// TIA Portal V19 export
// export: Created 2026-10-15T09:44:23.3519815Z, ExportSetting WithDefaults, DisplayName Totally Integrated Automation Portal, DisplayVersion V19, DisplayName TIA Portal Openness, DisplayVersion V19, DisplayName TIA Portal Version Control Interface, DisplayVersion V19, DisplayName STEP 7 Professional, DisplayVersion V19, DisplayName STEP 7 Safety, DisplayVersion V19, DisplayName WinCC Basic/Comfort/Advanced, DisplayVersion V19, DisplayName WinCC Unified, DisplayVersion V19
FUNCTION "ROLL_PB2" : Void   // FC14, SCL
{ S7_Optimized_Access := 'TRUE' }
VERSION : 0.1
// stored: AutoNumber true, IsIECCheckEnabled false, SetENOAutomatically false, UDAEnableTagReadback false
   VAR_TEMP
      r : Bool;
      a1 : Word;
      a2 : Word;
      activeDataBlock : Int;
      comparisonResults : Array[0..0] of Bool;
   END_VAR
BEGIN

   #r := FALSE;
   #a1 := W#16#0000;
   #a2 := W#16#0000;
   #activeDataBlock := 0;
   // PB2, STEP 5 network 1
   #r := ((NOT "ROLL_State".M[0, 1]) AND "ROLL_State".S5Timers[11].Q);
   "ROLL_State".M[4, 1] := #r;
   // PB2, STEP 5 network 2
   #r := ((NOT "ROLL_State".M[4, 1]) OR "ROLL_IO".Input[1, 0]);
   "ROLL_State".M[3, 1] := #r;
   // PB2, STEP 5 network 3
   #r := ((((NOT "ROLL_State".M[31, 4]) AND "ROLL_IO".Input[0, 4] AND "ROLL_State".M[4, 1]) OR "ROLL_State".M[31, 5]) AND "ROLL_IO".Input[0, 2]);
   "ROLL_State".M[4, 4] := #r;
   // PB2, STEP 5 network 4
   #r := (NOT "ROLL_IO".Input[11, 7]);
   IF #r THEN
       "ROLL_State".M[5, 0] := TRUE;
   END_IF;
   #r := "ROLL_State".M[3, 1];
   IF #r THEN
       "ROLL_State".M[5, 0] := FALSE;
   END_IF;
   // PB2, STEP 5 network 5
   #r := (NOT "ROLL_IO".Input[13, 5]);
   IF #r THEN
       "ROLL_State".M[5, 1] := TRUE;
   END_IF;
   #r := "ROLL_State".M[3, 1];
   IF #r THEN
       "ROLL_State".M[5, 1] := FALSE;
   END_IF;
   // PB2, STEP 5 network 6
   #r := (NOT "ROLL_IO".Input[13, 0]);
   IF #r THEN
       "ROLL_State".M[5, 2] := TRUE;
   END_IF;
   #r := "ROLL_State".M[3, 1];
   IF #r THEN
       "ROLL_State".M[5, 2] := FALSE;
   END_IF;
   // PB2, STEP 5 network 7
   #r := (NOT "ROLL_IO".Input[8, 5]);
   IF #r THEN
       "ROLL_State".M[5, 3] := TRUE;
   END_IF;
   #r := "ROLL_State".M[3, 1];
   IF #r THEN
       "ROLL_State".M[5, 3] := FALSE;
   END_IF;
   // PB2, STEP 5 network 8
   #r := "ROLL_State".M[0, 3];
   IF #r THEN
       "ROLL_State".M[5, 4] := TRUE;
   END_IF;
   #r := "ROLL_State".M[3, 1];
   IF #r THEN
       "ROLL_State".M[5, 4] := FALSE;
   END_IF;
   // PB2, STEP 5 network 9
   #r := "ROLL_State".M[0, 3];
   IF #r THEN
       "ROLL_State".M[5, 5] := TRUE;
   END_IF;
   #r := "ROLL_State".M[3, 1];
   IF #r THEN
       "ROLL_State".M[5, 5] := FALSE;
   END_IF;
   // PB2, STEP 5 network 10
   #r := "ROLL_IO".Input[3, 6];
   IF #r THEN
       "ROLL_State".M[5, 6] := TRUE;
   END_IF;
   #r := "ROLL_State".M[3, 1];
   IF #r THEN
       "ROLL_State".M[5, 6] := FALSE;
   END_IF;
   // PB2, STEP 5 network 11
   #r := (NOT "ROLL_IO".Input[3, 7]);
   IF #r THEN
       "ROLL_State".M[5, 7] := TRUE;
   END_IF;
   #r := "ROLL_State".M[3, 1];
   IF #r THEN
       "ROLL_State".M[5, 7] := FALSE;
   END_IF;
   // PB2, STEP 5 network 12
   #r := (NOT "ROLL_IO".Input[5, 2]);
   IF #r THEN
       "ROLL_State".M[6, 0] := TRUE;
   END_IF;
   #r := ("ROLL_IO".Input[5, 2] AND "ROLL_State".M[3, 1]);
   IF #r THEN
       "ROLL_State".M[6, 0] := FALSE;
   END_IF;
   // PB2, STEP 5 network 13
   #r := ((NOT "ROLL_IO".Input[5, 3]) AND "ROLL_State".S5Timers[31].Q);
   IF #r THEN
       "ROLL_State".M[6, 1] := TRUE;
   END_IF;
   #r := "ROLL_State".M[3, 1];
   IF #r THEN
       "ROLL_State".M[6, 1] := FALSE;
   END_IF;
   // PB2, STEP 5 network 14
   #r := (NOT "ROLL_IO".Input[5, 4]);
   IF #r THEN
       "ROLL_State".M[6, 2] := TRUE;
   END_IF;
   #r := ("ROLL_IO".Input[5, 4] AND "ROLL_State".M[3, 1]);
   IF #r THEN
       "ROLL_State".M[6, 2] := FALSE;
   END_IF;
   // PB2, STEP 5 network 15
   #r := ((NOT "ROLL_IO".Input[5, 5]) AND "ROLL_State".M[40, 5] AND "ROLL_State".S5Timers[17].Q);
   IF #r THEN
       "ROLL_State".M[6, 3] := TRUE;
   END_IF;
   #r := "ROLL_State".M[3, 1];
   IF #r THEN
       "ROLL_State".M[6, 3] := FALSE;
   END_IF;
   // PB2, STEP 5 network 16
   #r := ((NOT "ROLL_IO".Input[6, 0]) AND "ROLL_State".S5Timers[32].Q);
   IF #r THEN
       "ROLL_State".M[6, 4] := TRUE;
   END_IF;
   #r := "ROLL_State".M[3, 1];
   IF #r THEN
       "ROLL_State".M[6, 4] := FALSE;
   END_IF;
   // PB2, STEP 5 network 17
   #r := ((NOT "ROLL_IO".Input[6, 2]) AND "ROLL_State".S5Timers[33].Q);
   IF #r THEN
       "ROLL_State".M[6, 5] := TRUE;
   END_IF;
   #r := "ROLL_State".M[3, 1];
   IF #r THEN
       "ROLL_State".M[6, 5] := FALSE;
   END_IF;
   // PB2, STEP 5 network 18
   #r := "ROLL_State".M[0, 3];
   IF #r THEN
       "ROLL_State".M[6, 6] := TRUE;
   END_IF;
   #r := "ROLL_State".M[3, 1];
   IF #r THEN
       "ROLL_State".M[6, 6] := FALSE;
   END_IF;
   // PB2, STEP 5 network 19
   #r := ((NOT "ROLL_State".M[0, 3]) AND "ROLL_State".S5Timers[35].Q);
   IF #r THEN
       "ROLL_State".M[6, 7] := TRUE;
   END_IF;
   #r := "ROLL_State".M[3, 1];
   IF #r THEN
       "ROLL_State".M[6, 7] := FALSE;
   END_IF;
   // PB2, STEP 5 network 20
   #r := ((NOT "ROLL_State".M[0, 3]) AND "ROLL_State".S5Timers[36].Q);
   IF #r THEN
       "ROLL_State".M[7, 0] := TRUE;
   END_IF;
   #r := "ROLL_State".M[3, 1];
   IF #r THEN
       "ROLL_State".M[7, 0] := FALSE;
   END_IF;
   // PB2, STEP 5 network 21
   #r := ((NOT "ROLL_State".M[0, 3]) AND "ROLL_State".M[48, 1] AND "ROLL_State".S5Timers[37].Q);
   IF #r THEN
       "ROLL_State".M[7, 1] := TRUE;
   END_IF;
   #r := "ROLL_State".M[3, 1];
   IF #r THEN
       "ROLL_State".M[7, 1] := FALSE;
   END_IF;
   // PB2, STEP 5 network 22
   #r := ((NOT "ROLL_State".M[0, 3]) AND "ROLL_State".S5Timers[38].Q);
   IF #r THEN
       "ROLL_State".M[7, 2] := TRUE;
   END_IF;
   #r := "ROLL_State".M[3, 1];
   IF #r THEN
       "ROLL_State".M[7, 2] := FALSE;
   END_IF;
   // PB2, STEP 5 network 23
   #r := ((NOT "ROLL_IO".Input[5, 6]) AND "ROLL_State".S5Timers[16].Q);
   IF #r THEN
       "ROLL_State".M[7, 3] := TRUE;
   END_IF;
   #r := ("ROLL_IO".Input[5, 6] AND "ROLL_State".M[3, 1]);
   IF #r THEN
       "ROLL_State".M[7, 3] := FALSE;
   END_IF;
   // PB2, STEP 5 network 24
   #r := "ROLL_State".M[0, 3];
   IF #r THEN
       "ROLL_State".M[7, 4] := TRUE;
   END_IF;
   #r := "ROLL_State".M[3, 1];
   IF #r THEN
       "ROLL_State".M[7, 4] := FALSE;
   END_IF;
   // PB2, STEP 5 network 25
   #r := "ROLL_State".M[0, 3];
   IF #r THEN
       "ROLL_State".M[7, 5] := TRUE;
   END_IF;
   #r := "ROLL_State".M[3, 1];
   IF #r THEN
       "ROLL_State".M[7, 5] := FALSE;
   END_IF;
   // PB2, STEP 5 network 26
   #r := "ROLL_State".M[0, 3];
   IF #r THEN
       "ROLL_State".M[7, 6] := TRUE;
   END_IF;
   #r := "ROLL_State".M[3, 1];
   IF #r THEN
       "ROLL_State".M[7, 6] := FALSE;
   END_IF;
   // PB2, STEP 5 network 27
   #r := (NOT "ROLL_IO".Input[6, 7]);
   IF #r THEN
       "ROLL_State".M[7, 7] := TRUE;
   END_IF;
   #r := "ROLL_State".M[3, 1];
   IF #r THEN
       "ROLL_State".M[7, 7] := FALSE;
   END_IF;
   // PB2, STEP 5 network 28
   #a2 := #a1;
   #a1 := W#16#1050;
   #r := ((NOT "ROLL_IO".Input[7, 6]) AND "ROLL_IO".Output[20, 5]);
   "ROLL_TimerOp"(Number := 30,
                  Operation := 0,
                  Signal := #r,
                  Preset := #a1);
   #r := "ROLL_State".S5Timers[30].Q;
   IF #r THEN
       "ROLL_State".M[8, 6] := TRUE;
   END_IF;
   #r := "ROLL_State".M[3, 1];
   IF #r THEN
       "ROLL_State".M[8, 6] := FALSE;
   END_IF;
   // PB2, STEP 5 network 29
   #r := "ROLL_State".M[0, 3];
   IF #r THEN
       "ROLL_State".M[8, 7] := TRUE;
   END_IF;
   #r := "ROLL_State".M[3, 1];
   IF #r THEN
       "ROLL_State".M[8, 7] := FALSE;
   END_IF;
   // PB2, STEP 5 network 30
   #r := ((NOT "ROLL_IO".Input[13, 7]) AND "ROLL_State".M[4, 1]);
   IF #r THEN
       "ROLL_State".M[9, 0] := TRUE;
   END_IF;
   #r := ("ROLL_IO".Input[13, 7] AND "ROLL_State".M[3, 1]);
   IF #r THEN
       "ROLL_State".M[9, 0] := FALSE;
   END_IF;
   // PB2, STEP 5 network 31
   #r := "ROLL_State".M[0, 3];
   IF #r THEN
       "ROLL_State".M[9, 1] := TRUE;
   END_IF;
   #r := "ROLL_State".M[3, 1];
   IF #r THEN
       "ROLL_State".M[9, 1] := FALSE;
   END_IF;
   // PB2, STEP 5 network 32
   #r := ((NOT "ROLL_State".M[28, 4]) AND (NOT "ROLL_State".M[31, 5]) AND (((NOT "ROLL_State".M[20, 2]) AND ("ROLL_IO".Input[123, 5] OR "ROLL_IO".Input[123, 6])) OR "ROLL_State".M[70, 2] OR "ROLL_State".M[70, 3]) AND "ROLL_IO".Input[0, 4] AND "ROLL_State".M[4, 1]);
   IF #r THEN
       "ROLL_State".M[9, 2] := TRUE;
   END_IF;
   #r := "ROLL_State".M[3, 1];
   IF #r THEN
       "ROLL_State".M[9, 2] := FALSE;
   END_IF;
   // PB2, STEP 5 network 33
   #r := ("ROLL_State".M[4, 1] AND "ROLL_State".S5Timers[19].Q);
   IF #r THEN
       "ROLL_State".M[9, 3] := TRUE;
   END_IF;
   #r := "ROLL_State".M[3, 1];
   IF #r THEN
       "ROLL_State".M[9, 3] := FALSE;
   END_IF;
   // PB2, STEP 5 network 34
   #r := (((("ROLL_State".M[20, 4] OR "ROLL_State".M[20, 5]) AND "ROLL_IO".Input[0, 1] AND "ROLL_State".M[190, 6]) OR "ROLL_State".M[31, 5]) AND "ROLL_State".S5Timers[95].Q);
   "ROLL_State".M[9, 4] := #r;
   // PB2, STEP 5 network 35
   #r := "ROLL_State".M[0, 3];
   IF #r THEN
       "ROLL_State".M[9, 5] := TRUE;
   END_IF;
   #r := "ROLL_State".M[3, 1];
   IF #r THEN
       "ROLL_State".M[9, 5] := FALSE;
   END_IF;
   // PB2, STEP 5 network 36
   #r := "ROLL_State".M[0, 3];
   IF #r THEN
       "ROLL_State".M[9, 6] := TRUE;
   END_IF;
   #r := "ROLL_State".M[3, 1];
   IF #r THEN
       "ROLL_State".M[9, 6] := FALSE;
   END_IF;
   // PB2, STEP 5 network 37
   #r := "ROLL_State".M[0, 3];
   IF #r THEN
       "ROLL_State".M[9, 7] := TRUE;
   END_IF;
   #r := "ROLL_State".M[3, 1];
   IF #r THEN
       "ROLL_State".M[9, 7] := FALSE;
   END_IF;
   // PB2, STEP 5 network 38
   #r := ((NOT "ROLL_IO".Input[12, 0]) AND "ROLL_State".M[4, 1]);
   IF #r THEN
       "ROLL_State".M[10, 0] := TRUE;
   END_IF;
   #r := (((((NOT "ROLL_State".S5Timers[11].Q) AND "ROLL_IO".Input[3, 0]) OR "ROLL_IO".Input[12, 5]) AND "ROLL_State".M[3, 1]) OR (NOT "ROLL_State".M[4, 1]) OR "ROLL_State".M[0, 7]);
   IF #r THEN
       "ROLL_State".M[10, 0] := FALSE;
   END_IF;
   // PB2, STEP 5 network 39
   #r := ((NOT "ROLL_IO".Input[12, 6]) AND "ROLL_State".M[4, 1]);
   IF #r THEN
       "ROLL_State".M[10, 1] := TRUE;
   END_IF;
   #r := (((((NOT "ROLL_State".S5Timers[11].Q) AND "ROLL_IO".Input[3, 0]) OR "ROLL_IO".Input[12, 1]) AND "ROLL_State".M[3, 1]) OR (NOT "ROLL_State".M[4, 1]) OR "ROLL_State".M[0, 7]);
   IF #r THEN
       "ROLL_State".M[10, 1] := FALSE;
   END_IF;
   // PB2, STEP 5 network 40
   #r := "ROLL_State".M[0, 3];
   IF #r THEN
       "ROLL_State".M[10, 2] := TRUE;
   END_IF;
   #r := "ROLL_State".M[3, 1];
   IF #r THEN
       "ROLL_State".M[10, 2] := FALSE;
   END_IF;
   // PB2, STEP 5 network 41
   #r := "ROLL_State".M[0, 3];
   IF #r THEN
       "ROLL_State".M[10, 3] := TRUE;
   END_IF;
   #r := "ROLL_State".M[3, 1];
   IF #r THEN
       "ROLL_State".M[10, 3] := FALSE;
   END_IF;
   // PB2, STEP 5 network 42
   #r := "ROLL_State".M[0, 3];
   IF #r THEN
       "ROLL_State".M[10, 4] := TRUE;
   END_IF;
   #r := "ROLL_State".M[3, 1];
   IF #r THEN
       "ROLL_State".M[10, 4] := FALSE;
   END_IF;
   // PB2, STEP 5 network 43
   #r := "ROLL_State".M[0, 3];
   IF #r THEN
       "ROLL_State".M[10, 5] := TRUE;
   END_IF;
   #r := "ROLL_State".M[3, 1];
   IF #r THEN
       "ROLL_State".M[10, 5] := FALSE;
   END_IF;
   // PB2, STEP 5 network 44
   #r := "ROLL_State".M[0, 3];
   IF #r THEN
       "ROLL_State".M[10, 6] := TRUE;
   END_IF;
   #r := "ROLL_State".M[3, 1];
   IF #r THEN
       "ROLL_State".M[10, 6] := FALSE;
   END_IF;
   // PB2, STEP 5 network 45
   #r := "ROLL_State".M[0, 3];
   IF #r THEN
       "ROLL_State".M[10, 7] := TRUE;
   END_IF;
   #r := "ROLL_State".M[3, 1];
   IF #r THEN
       "ROLL_State".M[10, 7] := FALSE;
   END_IF;
   // PB2, STEP 5 network 46
   #r := ("ROLL_State".M[4, 1] AND "ROLL_State".M[63, 2]);
   IF #r THEN
       "ROLL_State".M[11, 0] := TRUE;
   END_IF;
   #r := "ROLL_State".M[3, 1];
   IF #r THEN
       "ROLL_State".M[11, 0] := FALSE;
   END_IF;
   // PB2, STEP 5 network 47
   #r := ("ROLL_IO".Input[13, 3] AND "ROLL_State".M[4, 1] AND "ROLL_State".S5Timers[112].Q);
   IF #r THEN
       "ROLL_State".M[11, 1] := TRUE;
   END_IF;
   #r := "ROLL_State".M[3, 1];
   IF #r THEN
       "ROLL_State".M[11, 1] := FALSE;
   END_IF;
   // PB2, STEP 5 network 48
   #r := ((NOT "ROLL_IO".Input[13, 3]) AND "ROLL_State".M[4, 1] AND "ROLL_State".S5Timers[15].Q);
   IF #r THEN
       "ROLL_State".M[11, 2] := TRUE;
   END_IF;
   #r := "ROLL_State".M[3, 1];
   IF #r THEN
       "ROLL_State".M[11, 2] := FALSE;
   END_IF;
   // PB2, STEP 5 network 49
   #r := ("ROLL_State".M[4, 1] AND "ROLL_State".M[63, 3]);
   IF #r THEN
       "ROLL_State".M[11, 3] := TRUE;
   END_IF;
   #r := "ROLL_State".M[3, 1];
   IF #r THEN
       "ROLL_State".M[11, 3] := FALSE;
   END_IF;
   // PB2, STEP 5 network 50
   #r := ("ROLL_State".M[190, 6] AND "ROLL_State".M[23, 2] AND "ROLL_State".M[60, 3]);
   IF #r THEN
       "ROLL_State".M[11, 4] := TRUE;
   END_IF;
   #r := "ROLL_State".M[3, 1];
   IF #r THEN
       "ROLL_State".M[11, 4] := FALSE;
   END_IF;
   // PB2, STEP 5 network 51
   #r := "ROLL_State".M[0, 3];
   IF #r THEN
       "ROLL_State".M[11, 5] := TRUE;
   END_IF;
   #r := "ROLL_State".M[3, 1];
   IF #r THEN
       "ROLL_State".M[11, 5] := FALSE;
   END_IF;
   // PB2, STEP 5 network 52
   #r := "ROLL_State".M[0, 3];
   IF #r THEN
       "ROLL_State".M[11, 6] := TRUE;
   END_IF;
   #r := "ROLL_State".M[3, 1];
   IF #r THEN
       "ROLL_State".M[11, 6] := FALSE;
   END_IF;
   // PB2, STEP 5 network 53
   #r := "ROLL_State".M[0, 3];
   IF #r THEN
       "ROLL_State".M[11, 7] := TRUE;
   END_IF;
   #r := "ROLL_State".M[3, 1];
   IF #r THEN
       "ROLL_State".M[11, 7] := FALSE;
   END_IF;
   // PB2, STEP 5 network 54
   #r := (NOT "ROLL_IO".Input[8, 3]);
   IF #r THEN
       "ROLL_State".M[12, 0] := TRUE;
   END_IF;
   #r := "ROLL_State".M[3, 1];
   IF #r THEN
       "ROLL_State".M[12, 0] := FALSE;
   END_IF;
   // PB2, STEP 5 network 55
   #r := ((NOT "ROLL_IO".Input[0, 7]) AND (NOT "ROLL_IO".Input[1, 4]) AND "ROLL_State".M[4, 4]);
   IF #r THEN
       "ROLL_State".M[12, 1] := TRUE;
   END_IF;
   #r := "ROLL_State".M[3, 1];
   IF #r THEN
       "ROLL_State".M[12, 1] := FALSE;
   END_IF;
   // PB2, STEP 5 network 56
   #r := "ROLL_State".M[0, 3];
   IF #r THEN
       "ROLL_State".M[12, 2] := TRUE;
   END_IF;
   #r := "ROLL_State".M[3, 1];
   IF #r THEN
       "ROLL_State".M[12, 2] := FALSE;
   END_IF;
   // PB2, STEP 5 network 57
   #r := "ROLL_State".M[0, 3];
   IF #r THEN
       "ROLL_State".M[12, 3] := TRUE;
   END_IF;
   #r := "ROLL_State".M[3, 1];
   IF #r THEN
       "ROLL_State".M[12, 3] := FALSE;
   END_IF;
   // PB2, STEP 5 network 58
   #r := "ROLL_State".M[0, 3];
   IF #r THEN
       "ROLL_State".M[13, 0] := TRUE;
   END_IF;
   #r := "ROLL_State".M[3, 1];
   IF #r THEN
       "ROLL_State".M[13, 0] := FALSE;
   END_IF;
   // PB2, STEP 5 network 59
   #r := (NOT "ROLL_IO".Input[3, 2]);
   IF #r THEN
       "ROLL_State".M[13, 1] := TRUE;
   END_IF;
   #r := "ROLL_State".M[3, 1];
   IF #r THEN
       "ROLL_State".M[13, 1] := FALSE;
   END_IF;
   // PB2, STEP 5 network 60
   #r := ((NOT "ROLL_IO".Input[4, 7]) AND "ROLL_IO".Input[0, 1] AND "ROLL_State".M[190, 6] AND "ROLL_State".M[27, 4]);
   IF #r THEN
       "ROLL_State".M[13, 2] := TRUE;
   END_IF;
   #r := "ROLL_State".M[3, 1];
   IF #r THEN
       "ROLL_State".M[13, 2] := FALSE;
   END_IF;
   // PB2, STEP 5 network 61
   #r := (NOT "ROLL_IO".Input[5, 0]);
   IF #r THEN
       "ROLL_State".M[13, 3] := TRUE;
   END_IF;
   #r := ("ROLL_IO".Input[5, 0] AND "ROLL_State".M[3, 1]);
   IF #r THEN
       "ROLL_State".M[13, 3] := FALSE;
   END_IF;
   // PB2, STEP 5 network 62
   #r := (NOT "ROLL_IO".Input[10, 7]);
   IF #r THEN
       "ROLL_State".M[13, 4] := TRUE;
   END_IF;
   #r := ("ROLL_IO".Input[10, 7] AND "ROLL_State".M[3, 1]);
   IF #r THEN
       "ROLL_State".M[13, 4] := FALSE;
   END_IF;
   // PB2, STEP 5 network 63
   #r := (NOT "ROLL_IO".Input[4, 5]);
   IF #r THEN
       "ROLL_State".M[13, 7] := TRUE;
   END_IF;
   #r := "ROLL_State".M[3, 1];
   IF #r THEN
       "ROLL_State".M[13, 7] := FALSE;
   END_IF;
   // PB2, STEP 5 network 64
   #a2 := #a1;
   #a1 := W#16#2020;
   #r := (((NOT "ROLL_IO".Input[10, 0]) OR (NOT "ROLL_IO".Input[10, 1]) OR (NOT "ROLL_IO".Input[10, 2]) OR (NOT "ROLL_IO".Input[10, 3])) AND "ROLL_IO".Output[19, 1]);
   "ROLL_TimerOp"(Number := 50,
                  Operation := 0,
                  Signal := #r,
                  Preset := #a1);
   // PB2, STEP 5 network 65
   #r := ((NOT "ROLL_IO".Input[10, 0]) AND "ROLL_State".S5Timers[50].Q);
   IF #r THEN
       "ROLL_State".M[14, 0] := TRUE;
   END_IF;
   #r := "ROLL_State".M[3, 1];
   IF #r THEN
       "ROLL_State".M[14, 0] := FALSE;
   END_IF;
   // PB2, STEP 5 network 66
   #r := ((NOT "ROLL_IO".Input[10, 1]) AND "ROLL_State".S5Timers[50].Q);
   IF #r THEN
       "ROLL_State".M[14, 1] := TRUE;
   END_IF;
   #r := "ROLL_State".M[3, 1];
   IF #r THEN
       "ROLL_State".M[14, 1] := FALSE;
   END_IF;
   // PB2, STEP 5 network 67
   #r := ((NOT "ROLL_IO".Input[10, 2]) AND "ROLL_State".S5Timers[50].Q);
   IF #r THEN
       "ROLL_State".M[14, 2] := TRUE;
   END_IF;
   #r := "ROLL_State".M[3, 1];
   IF #r THEN
       "ROLL_State".M[14, 2] := FALSE;
   END_IF;
   // PB2, STEP 5 network 68
   #r := ((NOT "ROLL_IO".Input[10, 3]) AND "ROLL_State".S5Timers[50].Q);
   IF #r THEN
       "ROLL_State".M[14, 3] := TRUE;
   END_IF;
   #r := "ROLL_State".M[3, 1];
   IF #r THEN
       "ROLL_State".M[14, 3] := FALSE;
   END_IF;
   // PB2, STEP 5 network 69
   #r := "ROLL_State".M[0, 3];
   IF #r THEN
       "ROLL_State".M[15, 2] := TRUE;
   END_IF;
   #r := "ROLL_State".M[3, 1];
   IF #r THEN
       "ROLL_State".M[15, 2] := FALSE;
   END_IF;
   // PB2, STEP 5 network 70
   #r := "ROLL_State".M[0, 3];
   IF #r THEN
       "ROLL_State".M[15, 3] := TRUE;
   END_IF;
   #r := "ROLL_State".M[3, 1];
   IF #r THEN
       "ROLL_State".M[15, 3] := FALSE;
   END_IF;
   // PB2, STEP 5 network 71
   #r := "ROLL_State".M[0, 3];
   IF #r THEN
       "ROLL_State".M[15, 4] := TRUE;
   END_IF;
   #r := "ROLL_State".M[3, 1];
   IF #r THEN
       "ROLL_State".M[15, 4] := FALSE;
   END_IF;
   // PB2, STEP 5 network 72
   #r := (NOT "ROLL_IO".Input[4, 0]);
   IF #r THEN
       "ROLL_State".M[15, 5] := TRUE;
   END_IF;
   #r := "ROLL_State".M[3, 1];
   IF #r THEN
       "ROLL_State".M[15, 5] := FALSE;
   END_IF;
   // PB2, STEP 5 network 73
   #r := (NOT "ROLL_IO".Input[4, 1]);
   IF #r THEN
       "ROLL_State".M[15, 6] := TRUE;
   END_IF;
   #r := "ROLL_State".M[3, 1];
   IF #r THEN
       "ROLL_State".M[15, 6] := FALSE;
   END_IF;
   // PB2, STEP 5 network 74
   #r := (NOT "ROLL_IO".Input[4, 2]);
   IF #r THEN
       "ROLL_State".M[15, 7] := TRUE;
   END_IF;
   #r := "ROLL_State".M[3, 1];
   IF #r THEN
       "ROLL_State".M[15, 7] := FALSE;
   END_IF;
   // PB2, STEP 5 network 75
   #r := "ROLL_State".M[16, 0];
   IF #r THEN
       "ROLL_State".M[16, 0] := TRUE;
   END_IF;
   #r := "ROLL_State".M[3, 1];
   IF #r THEN
       "ROLL_State".M[16, 0] := FALSE;
   END_IF;
   // PB2, STEP 5 network 76
   #r := "ROLL_State".M[16, 1];
   IF #r THEN
       "ROLL_State".M[16, 1] := TRUE;
   END_IF;
   #r := "ROLL_State".M[3, 1];
   IF #r THEN
       "ROLL_State".M[16, 1] := FALSE;
   END_IF;
   // PB2, STEP 5 network 77
   #r := "ROLL_State".M[16, 2];
   IF #r THEN
       "ROLL_State".M[16, 2] := TRUE;
   END_IF;
   #r := "ROLL_State".M[3, 1];
   IF #r THEN
       "ROLL_State".M[16, 2] := FALSE;
   END_IF;
   // PB2, STEP 5 network 78
   #r := ("ROLL_State".M[34, 1] AND "ROLL_State".M[4, 1]);
   IF #r THEN
       "ROLL_State".M[16, 3] := TRUE;
   END_IF;
   #r := "ROLL_State".M[3, 1];
   IF #r THEN
       "ROLL_State".M[16, 3] := FALSE;
   END_IF;
   // PB2, STEP 5 network 79
   #r := "ROLL_State".M[16, 4];
   IF #r THEN
       "ROLL_State".M[16, 4] := TRUE;
   END_IF;
   #r := ((NOT "ROLL_IO".Input[123, 1]) AND (NOT "ROLL_IO".Input[123, 4]) AND (NOT "ROLL_IO".Input[123, 5]) AND (NOT "ROLL_IO".Input[123, 6]) AND (NOT "ROLL_IO".Input[125, 0]) AND (NOT "ROLL_IO".Input[125, 1]) AND "ROLL_State".M[3, 1]);
   IF #r THEN
       "ROLL_State".M[16, 4] := FALSE;
   END_IF;
   // PB2, STEP 5 network 80
   #r := "ROLL_State".M[16, 5];
   IF #r THEN
       "ROLL_State".M[16, 5] := TRUE;
   END_IF;
   #r := "ROLL_State".M[3, 1];
   IF #r THEN
       "ROLL_State".M[16, 5] := FALSE;
   END_IF;
   // PB2, STEP 5 network 81
   #r := ((NOT "ROLL_IO".Input[3, 4]) AND "ROLL_State".M[4, 1]);
   IF #r THEN
       "ROLL_State".M[16, 6] := TRUE;
   END_IF;
   #r := ("ROLL_IO".Input[3, 4] AND "ROLL_State".M[3, 1]);
   IF #r THEN
       "ROLL_State".M[16, 6] := FALSE;
   END_IF;
   // PB2, STEP 5 network 82
   #r := ((NOT "ROLL_IO".Input[3, 1]) AND ((("ROLL_State".M[190, 5] OR "ROLL_State".M[190, 6]) AND "ROLL_IO".Input[0, 1]) OR "ROLL_State".M[4, 4]) AND "ROLL_State".M[4, 1]);
   IF #r THEN
       "ROLL_State".M[16, 7] := TRUE;
   END_IF;
   #r := "ROLL_State".M[3, 1];
   IF #r THEN
       "ROLL_State".M[16, 7] := FALSE;
   END_IF;
   // PB2, STEP 5 network 83
   #r := ((NOT "ROLL_IO".Input[3, 5]) AND "ROLL_State".M[4, 1]);
   IF #r THEN
       "ROLL_State".M[17, 0] := TRUE;
   END_IF;
   #r := ("ROLL_IO".Input[3, 5] AND "ROLL_State".M[3, 1]);
   IF #r THEN
       "ROLL_State".M[17, 0] := FALSE;
   END_IF;
   // PB2, STEP 5 network 84
   #r := "ROLL_State".M[0, 3];
   IF #r THEN
       "ROLL_State".M[17, 1] := TRUE;
   END_IF;
   #r := "ROLL_State".M[3, 1];
   IF #r THEN
       "ROLL_State".M[17, 1] := FALSE;
   END_IF;
   // PB2, STEP 5 network 85
   #r := "ROLL_State".M[0, 3];
   IF #r THEN
       "ROLL_State".M[17, 2] := TRUE;
   END_IF;
   #r := "ROLL_State".M[3, 1];
   IF #r THEN
       "ROLL_State".M[17, 2] := FALSE;
   END_IF;
   // PB2, STEP 5 network 86
   #r := "ROLL_State".M[0, 3];
   IF #r THEN
       "ROLL_State".M[17, 3] := TRUE;
   END_IF;
   #r := "ROLL_State".M[3, 1];
   IF #r THEN
       "ROLL_State".M[17, 3] := FALSE;
   END_IF;
   // PB2, STEP 5 network 87
   #r := "ROLL_State".M[0, 3];
   IF #r THEN
       "ROLL_State".M[17, 4] := TRUE;
   END_IF;
   #r := "ROLL_State".M[3, 1];
   IF #r THEN
       "ROLL_State".M[17, 4] := FALSE;
   END_IF;
   // PB2, STEP 5 network 88
   #r := "ROLL_State".M[0, 3];
   IF #r THEN
       "ROLL_State".M[17, 5] := TRUE;
   END_IF;
   #r := "ROLL_State".M[3, 1];
   IF #r THEN
       "ROLL_State".M[17, 5] := FALSE;
   END_IF;
   // PB2, STEP 5 network 89
   #r := "ROLL_State".M[0, 3];
   IF #r THEN
       "ROLL_State".M[17, 6] := TRUE;
   END_IF;
   #r := "ROLL_State".M[3, 1];
   IF #r THEN
       "ROLL_State".M[17, 6] := FALSE;
   END_IF;
   // PB2, STEP 5 network 90
   #r := "ROLL_State".M[0, 3];
   IF #r THEN
       "ROLL_State".M[17, 7] := TRUE;
   END_IF;
   #r := "ROLL_State".M[3, 1];
   IF #r THEN
       "ROLL_State".M[17, 7] := FALSE;
   END_IF;
   // PB2, STEP 5 network 91
   #r := "ROLL_State".M[0, 3];
   IF #r THEN
       "ROLL_State".M[18, 0] := TRUE;
   END_IF;
   #r := "ROLL_State".M[3, 1];
   IF #r THEN
       "ROLL_State".M[18, 0] := FALSE;
   END_IF;
   // PB2, STEP 5 network 92
   #r := ((NOT "ROLL_IO".Input[14, 0]) AND ((("ROLL_State".M[190, 5] OR "ROLL_State".M[190, 6]) AND ("ROLL_State".M[23, 0] OR "ROLL_State".M[23, 1] OR "ROLL_State".M[23, 2] OR "ROLL_State".M[23, 3])) OR ("ROLL_State".M[16, 3] AND "ROLL_State".M[31, 4] AND "ROLL_State".M[37, 2]) OR "ROLL_State".M[74, 0]));
   IF #r THEN
       "ROLL_State".M[18, 1] := TRUE;
   END_IF;
   #r := "ROLL_State".M[3, 1];
   IF #r THEN
       "ROLL_State".M[18, 1] := FALSE;
   END_IF;
   // PB2, STEP 5 network 93
   #r := "ROLL_State".M[0, 3];
   IF #r THEN
       "ROLL_State".M[18, 2] := TRUE;
   END_IF;
   #r := "ROLL_State".M[3, 1];
   IF #r THEN
       "ROLL_State".M[18, 2] := FALSE;
   END_IF;
   // PB2, STEP 5 network 94
   #r := "ROLL_State".M[0, 3];
   IF #r THEN
       "ROLL_State".M[18, 3] := TRUE;
   END_IF;
   #r := "ROLL_State".M[3, 1];
   IF #r THEN
       "ROLL_State".M[18, 3] := FALSE;
   END_IF;
   // PB2, STEP 5 network 95
   #r := "ROLL_State".M[0, 3];
   IF #r THEN
       "ROLL_State".M[18, 4] := TRUE;
   END_IF;
   #r := "ROLL_State".M[3, 1];
   IF #r THEN
       "ROLL_State".M[18, 4] := FALSE;
   END_IF;
   // PB2, STEP 5 network 96
   #r := "ROLL_State".M[0, 3];
   IF #r THEN
       "ROLL_State".M[18, 5] := TRUE;
   END_IF;
   #r := "ROLL_State".M[3, 1];
   IF #r THEN
       "ROLL_State".M[18, 5] := FALSE;
   END_IF;
   // PB2, STEP 5 network 97
   #r := "ROLL_State".M[0, 3];
   IF #r THEN
       "ROLL_State".M[18, 6] := TRUE;
   END_IF;
   #r := "ROLL_State".M[3, 1];
   IF #r THEN
       "ROLL_State".M[18, 6] := FALSE;
   END_IF;
   // PB2, STEP 5 network 98
   #r := "ROLL_State".M[0, 3];
   IF #r THEN
       "ROLL_State".M[18, 7] := TRUE;
   END_IF;
   #r := "ROLL_State".M[3, 1];
   IF #r THEN
       "ROLL_State".M[18, 7] := FALSE;
   END_IF;
   // PB2, STEP 5 network 99
   #r := "ROLL_State".M[0, 3];
   IF #r THEN
       "ROLL_State".M[19, 0] := TRUE;
   END_IF;
   #r := "ROLL_State".M[3, 1];
   IF #r THEN
       "ROLL_State".M[19, 0] := FALSE;
   END_IF;
   // PB2, STEP 5 network 100
   #r := "ROLL_State".M[0, 3];
   IF #r THEN
       "ROLL_State".M[19, 1] := TRUE;
   END_IF;
   #r := "ROLL_State".M[3, 1];
   IF #r THEN
       "ROLL_State".M[19, 1] := FALSE;
   END_IF;
   // PB2, STEP 5 network 101
   #r := "ROLL_State".M[0, 3];
   IF #r THEN
       "ROLL_State".M[19, 2] := TRUE;
   END_IF;
   #r := "ROLL_State".M[3, 1];
   IF #r THEN
       "ROLL_State".M[19, 2] := FALSE;
   END_IF;
   // PB2, STEP 5 network 102
   #r := "ROLL_State".M[0, 3];
   IF #r THEN
       "ROLL_State".M[19, 3] := TRUE;
   END_IF;
   #r := "ROLL_State".M[3, 1];
   IF #r THEN
       "ROLL_State".M[19, 3] := FALSE;
   END_IF;
   // PB2, STEP 5 network 103
   #r := "ROLL_State".M[0, 3];
   IF #r THEN
       "ROLL_State".M[19, 4] := TRUE;
   END_IF;
   #r := "ROLL_State".M[3, 1];
   IF #r THEN
       "ROLL_State".M[19, 4] := FALSE;
   END_IF;
   // PB2, STEP 5 network 104
   #r := "ROLL_State".M[0, 3];
   IF #r THEN
       "ROLL_State".M[19, 5] := TRUE;
   END_IF;
   #r := "ROLL_State".M[3, 1];
   IF #r THEN
       "ROLL_State".M[19, 5] := FALSE;
   END_IF;
   // PB2, STEP 5 network 105
   #r := "ROLL_State".M[0, 3];
   IF #r THEN
       "ROLL_State".M[19, 6] := TRUE;
   END_IF;
   #r := "ROLL_State".M[3, 1];
   IF #r THEN
       "ROLL_State".M[19, 6] := FALSE;
   END_IF;
   // PB2, STEP 5 network 106
   #r := "ROLL_State".M[0, 3];
   IF #r THEN
       "ROLL_State".M[19, 7] := TRUE;
   END_IF;
   #r := "ROLL_State".M[3, 1];
   IF #r THEN
       "ROLL_State".M[19, 7] := FALSE;
   END_IF;
   // PB2, STEP 5 network 107
   RETURN;
END_FUNCTION
